(* IEC 61131-3 sources: plc-iiot-stack/tests/POUs/FB_MqttDiag_Test, 13 files *)

(* ---- BackoffDoublesUpToMaximum.method.decl.st ---- *)
// Пауза между попытками: 1, 2, 4 с и дальше 4 с (tBackoffMax).
METHOD PRIVATE BackoffDoublesUpToMaximum
VAR_INST
    fbFake : FB_MqttClientFake;
    fbDiag : FB_MqttDiag;
    stCfg : ST_MqttBrokerCfg;
END_VAR

(* ---- BirthRefusedMeansNotReady.method.decl.st ---- *)
// Рождение не принято клиентом — связь есть, но публиковать нельзя; повтор.
METHOD PRIVATE BirthRefusedMeansNotReady
VAR_INST
    fbFake : FB_MqttClientFake;
    fbDiag : FB_MqttDiag;
    stCfg : ST_MqttBrokerCfg;
END_VAR

(* ---- ConnectionLossCountsAndReconnects.method.decl.st ---- *)
// Потеря связи: разрыв, код -4, пауза 1 с, переподключение и новое рождение.
METHOD PRIVATE ConnectionLossCountsAndReconnects
VAR_INST
    fbFake : FB_MqttClientFake;
    fbDiag : FB_MqttDiag;
    stCfg : ST_MqttBrokerCfg;
END_VAR

(* ---- ConnectSetsLwtAndPublishesBirth.method.decl.st ---- *)
// Подключение: завещание offline/lwt, рождение online/birth (QoS 1, retain), xReady.
METHOD PRIVATE ConnectSetsLwtAndPublishesBirth
VAR_INST
    fbFake : FB_MqttClientFake;
    fbDiag : FB_MqttDiag;
    stCfg : ST_MqttBrokerCfg;
END_VAR

VAR
    uiIdx : UINT;
END_VAR

(* ---- ConnectSetsLwtAndPublishesBirth.method.impl.st ---- *)
coUnit.TEST('ConnectSetsLwtAndPublishesBirth');

fbDiag(xEnable := TRUE, itfClient := fbFake, ltNow := LTIME#1H, uliTs_ms := 1792137600250,
    sTopicPrefix := 'vodokanal/kns1/station',
       stBroker := stCfg);

AssertTrue(Condition := fbDiag.eState = E_MqttConnState.Connected, Message := 'connected in the same call');
AssertTrue(Condition := fbDiag.xReady AND fbDiag.eNe107 = E_IiotNe107.Good, Message := 'ready, NE107 Good');
AssertEquals_STRING(Expected := 'vodokanal/kns1/station/PLC1/status/connection', Actual := fbFake.stLastCfg.sWillTopic,
    Message := 'LWT topic');
AssertEquals_STRING(
    Expected := '{"schema_version":"1.1","ts":1792137600250,"node":"PLC1","state":"offline","reason":"lwt"}',
    Actual := fbFake.stLastCfg.sWillPayload, Message := 'LWT payload');
AssertTrue(Condition := fbFake.stLastCfg.xWillRetain, Message := 'LWT retained');
AssertEquals_STRING(Expected := CONCAT('{"schema_version":"1.1","ts":1792137600250,"node":"PLC1","state":"online",',
    '"reason":"birth","source":"codesys","sw_version":"0.1.0","period_ms":60000}'),
    Actual := fbFake.LastPayload(sTopic := 'vodokanal/kns1/station/PLC1/status/connection'),
        Message := 'birth payload');
uiIdx := fbFake.FindLast(sTopic := 'vodokanal/kns1/station/PLC1/status/connection');
AssertTrue(Condition := uiIdx > 0, Message := 'birth published');
IF uiIdx > 0 THEN
    AssertTrue(Condition := fbFake.aPub[uiIdx].xRetain AND fbFake.aPub[uiIdx].eQos = E_MqttQos.AtLeastOnce,
               Message := 'birth: QoS 1, retain');
END_IF

coUnit.TEST_FINISHED();

(* ---- ConnectTimeoutGoesToBackoff.method.decl.st ---- *)
// Нет CONNACK за tConnectTimeout — неудача, код -2, разрыв, пауза, статус S.
METHOD PRIVATE ConnectTimeoutGoesToBackoff
VAR_INST
    fbFake : FB_MqttClientFake;
    fbDiag : FB_MqttDiag;
    stCfg : ST_MqttBrokerCfg;
END_VAR

(* ---- DegradedWhenPublishFailuresGrow.method.decl.st ---- *)
// Рост отказов публикаций за окно — M; нет роста — снова Good.
METHOD PRIVATE DegradedWhenPublishFailuresGrow
VAR_INST
    fbFake : FB_MqttClientFake;
    fbDiag : FB_MqttDiag;
    stCfg : ST_MqttBrokerCfg;
END_VAR

(* ---- DisabledIsCheckFunctionWithoutConnect.method.decl.st ---- *)
// Выключено: Disabled, статус C, подключений нет.
METHOD PRIVATE DisabledIsCheckFunctionWithoutConnect
VAR_INST
    fbFake : FB_MqttClientFake;
    fbDiag : FB_MqttDiag;
    stCfg : ST_MqttBrokerCfg;
END_VAR

(* ---- DisableWhileConnectedPublishesShutdown.method.decl.st ---- *)
// Выключение при связи: offline/shutdown, затем разрыв в следующем вызове.
METHOD PRIVATE DisableWhileConnectedPublishesShutdown
VAR_INST
    fbFake : FB_MqttClientFake;
    fbDiag : FB_MqttDiag;
    stCfg : ST_MqttBrokerCfg;
END_VAR

(* ---- FailureAfterThresholdAndResetAfterStableLink.method.decl.st ---- *)
// Три неудачи подряд — F; после tStable связи счётчик и пауза сбрасываются.
METHOD PRIVATE FailureAfterThresholdAndResetAfterStableLink
VAR_INST
    fbFake : FB_MqttClientFake;
    fbDiag : FB_MqttDiag;
    stCfg : ST_MqttBrokerCfg;
END_VAR

(* ---- NoClockNoConnect.method.decl.st ---- *)
// Часы ПЛК не установлены: подключения нет, код -5, статус C.
METHOD PRIVATE NoClockNoConnect
VAR_INST
    fbFake : FB_MqttClientFake;
    fbDiag : FB_MqttDiag;
    stCfg : ST_MqttBrokerCfg;
END_VAR

(* ---- RejectedConnectUsesClientErrorCode.method.decl.st ---- *)
// Connect() отклонён: код ошибки клиента, без него — -3.
METHOD PRIVATE RejectedConnectUsesClientErrorCode
VAR_INST
    fbFake : FB_MqttClientFake;
    fbDiag : FB_MqttDiag;
    stCfg : ST_MqttBrokerCfg;
END_VAR

(* ---- TimeGoingBackwardsRestartsTimeout.method.decl.st ---- *)
// Время пошло назад — отсчёт тайм-аута заново, без зависания.
METHOD PRIVATE TimeGoingBackwardsRestartsTimeout
VAR_INST
    fbFake : FB_MqttClientFake;
    fbDiag : FB_MqttDiag;
    stCfg : ST_MqttBrokerCfg;
END_VAR
